Fanuc KAREL source: KT00704.KL

PROGRAM KT00704
%NOLOCKGROUP
VAR
  C1: CONFIG
  C2: CONFIG
  OUT: REAL
BEGIN
  C1.CFG_FLIP = TRUE
  C2.CFG_FLIP = FALSE
  C1.CFG_FLIP = TRUE
  C2.CFG_FLIP = FALSE
  OUT = - C1
END KT00704
